Fanuc KAREL source: KC00019.KL

PROGRAM KC00019
%NOLOCKGROUP
VAR
  I: INTEGER
  J: INTEGER
  K: INTEGER
  R: REAL
  B: BOOLEAN
  S: STRING[80]
  T: STRING[80]
  P: PATH
  Q: PATH
  AI: ARRAY[8] OF INTEGER
  AB: ARRAY[244] OF BYTE
  F: FILE
  SA: ARRAY[8] OF STRING[80]
  SB: ARRAY[8] OF STRING[80]
BEGIN
  XML_GETDATA(F,I,SA,SB,S,B,J)
END KC00019
